// TwinCAT 3 PLC project TcoAteqMeasurementTests
// Title: TcoAteqMeasurementTests
// Company: Vortex.Library
// ProjectVersion: 0.6.0.913
// ProgramVersion: 3.1.4024.12
// libraries:
//   TcoAteqMeasurement, 0.6.0.913 (Vortex.Library)
//   Tc2_Standard, * (Beckhoff Automation GmbH)
//   Tc2_System, * (Beckhoff Automation GmbH)
//   Tc3_Module, * (Beckhoff Automation GmbH)
//   TcoIo, 0.6.0.913 (Vortex.Library)
//   TcoCore, 0.6.0.913 (Vortex.Library)
// project tree:
//   GVLs/ GVL.TcGVL
//   / PlcTask.TcTTO
//   POUs/ MAIN.TcPOU
//   Tests/TcoAteqG6/ eTcoAteqG6Tests.TcDUT, TcoAteqG6Simulator.TcPOU, TcoAteqG6TestContext.TcPOU
//   Tests/TcoContext/ WpfContext.TcPOU
// (motion and I/O tree: see PLC project tcoateqmeasurement)
// real-time tasks:
//   TASK PlcTask: cycle T#10ms, priority 20, ADS port 350
//   TASK PlcTask1: cycle T#10ms, priority 21, ADS port 351

CONFIGURATION TcoAteqMeasurementTests
    RESOURCE PLC ON TwinCAT3
        TASK PlcTask(INTERVAL := T#10ms, PRIORITY := 21);
        PROGRAM MAIN WITH PlcTask : MAIN;
    END_RESOURCE
END_CONFIGURATION

// ---- Tests/TcoAteqG6/eTcoAteqG6Tests.TcDUT
{attribute 'qualified_only'}
{attribute 'strict'}
TYPE eTcoAteqG6Tests :
(
	None := 0,
	Restore := 10,
	Run := 20,
	Reset := 30,
	SelectProgram := 40,
	StartCycle := 50,
	ReadLastResult := 60,
	SpecialCycle := 70,
	ReadParameters := 80,
	ReadPresetParameters := 90,
	ReadParameter := 100,
	InvokeStartCycle := 110,
	InvokeSelectProgram := 120,
	InvokeReset := 130
);
END_TYPE

// ---- GVLs/GVL.TcGVL
{attribute 'qualified_only'}
VAR_GLOBAL
	Ateq1 : TcoAteqMeasurement.TcoAteqG6Pn_IO_v_3_5_x;
END_VAR

// ---- POUs/MAIN.TcPOU
PROGRAM MAIN
VAR
	_g6TestContext : TcoAteqG6TestContext;

	_wpfContext : WpfContext;
	_wpfContextCall : BOOL := FALSE;
END_VAR

_g6TestContext.ProbeRun();

IF _wpfContextCall THEN
	_wpfContext.Run();
END_IF

END_PROGRAM

// ---- Tests/TcoAteqG6/TcoAteqG6TestContext.TcPOU
(*~
	<docu>
		<summary>
			Test context of TcoAteqG6Pn_v_3_5_x. _inImage is the input image of the instrument: written by the simulator
			when _simulate = TRUE, otherwise directly by the test. _outImage is what the component put on the wire.
		</summary>
	</docu>
~*)
FUNCTION_BLOCK TcoAteqG6TestContext EXTENDS TcoCore._internals_TcoContext
VAR
	_sut : TcoAteqMeasurement.TcoAteqG6Pn_v_3_5_x(THIS^);
	_io : TcoAteqMeasurement.TcoAteqG6Pn_IO_v_3_5_x;
	_sim : TcoAteqG6Simulator;
	_simulate : BOOL;
	_inImage : ARRAY[0..255] OF BYTE;
	_outImage : ARRAY[0..255] OF BYTE;
	_program : INT;
	_specialCycle : TcoAteqMeasurement.eTcoAteqG6_SpecialCycle_v_3_5_x;
	_instruction : BYTE;
	_parameter : TcoAteqMeasurement.eTcoAteqG6_ParameterId_v_3_5_x;
	_request : TcoAteqMeasurement.TcoAteqG6_ParameterRequest_v_3_5_x;
	_taskDone : BOOL;
	_taskError : BOOL;
	_startCycleBusy : BOOL;
	_selectProgramBusy : BOOL;
	_resetBusy : BOOL;
END_VAR
VAR
	{attribute 'hide'}
	_i : INT;
END_VAR

METHOD PROTECTED Main
//*************INSTRUMENT SIMULATOR*******
IF _simulate THEN
	_sim.Step(inoOut := _outImage, inoIn := _inImage);
END_IF

//*************INPUT IMAGE****************
MEMCPY(destAddr := ADR(_io.In.In1), srcAddr := ADR(_inImage[0]), n := 64);
MEMCPY(destAddr := ADR(_io.In.In2), srcAddr := ADR(_inImage[64]), n := 64);
MEMCPY(destAddr := ADR(_io.In.In3), srcAddr := ADR(_inImage[128]), n := 64);
MEMCPY(destAddr := ADR(_io.In.In4), srcAddr := ADR(_inImage[192]), n := 64);

CASE _testId OF
	eTcoAteqG6Tests.Restore:
		_sut.Restore();
		_sut._messenger.Clear();
		_sim.Reset();
		FOR _i := 0 TO 255 DO
			_inImage[_i] := 0;
		END_FOR
		_taskDone := FALSE;
		_taskError := FALSE;
		ProbeDoneWhen(TRUE);
	eTcoAteqG6Tests.Run:
		;
	eTcoAteqG6Tests.Reset:
		_taskDone := _sut.Reset().Done;
		_taskError := _sut.ResetTask.Error;
		ProbeDoneWhen(_taskDone OR _taskError);
	eTcoAteqG6Tests.SelectProgram:
		_taskDone := _sut.SelectProgram(_program).Done;
		_taskError := _sut.SelectProgramTask.Error;
		ProbeDoneWhen(_taskDone OR _taskError);
	eTcoAteqG6Tests.StartCycle:
		_taskDone := _sut.StartCycle(_program).Done;
		_taskError := _sut.StartCycleTask.Error;
		ProbeDoneWhen(_taskDone OR _taskError);
	eTcoAteqG6Tests.ReadLastResult:
		_taskDone := _sut.ReadLastResult().Done;
		_taskError := _sut.ReadLastResultTask.Error;
		ProbeDoneWhen(_taskDone OR _taskError);
	eTcoAteqG6Tests.SpecialCycle:
		_taskDone := _sut.SpecialCycle(_specialCycle, _instruction).Done;
		_taskError := _sut.SpecialCycleTask.Error;
		ProbeDoneWhen(_taskDone OR _taskError);
	eTcoAteqG6Tests.ReadParameters:
		_taskDone := _sut.ReadParameters(_request).Done;
		_taskError := _sut.ReadParametersTask.Error;
		ProbeDoneWhen(_taskDone OR _taskError);
	eTcoAteqG6Tests.ReadPresetParameters:
		_taskDone := _sut.ReadPresetParameters().Done;
		_taskError := _sut.ReadParametersTask.Error;
		ProbeDoneWhen(_taskDone OR _taskError);
	eTcoAteqG6Tests.ReadParameter:
		_taskDone := _sut.ReadParameter(_parameter).Done;
		_taskError := _sut.ReadParametersTask.Error;
		ProbeDoneWhen(_taskDone OR _taskError);
	eTcoAteqG6Tests.InvokeStartCycle:
		_sut.StartCycle(_program);
		ProbeDoneWhen(TRUE);
	eTcoAteqG6Tests.InvokeSelectProgram:
		_sut.SelectProgram(_program);
		ProbeDoneWhen(TRUE);
	eTcoAteqG6Tests.InvokeReset:
		_sut.Reset();
		ProbeDoneWhen(TRUE);
END_CASE

_sut(inoData := _io);

//*************OUTPUT IMAGE***************
MEMCPY(destAddr := ADR(_outImage[0]), srcAddr := ADR(_io.Out.Out1), n := 64);
MEMCPY(destAddr := ADR(_outImage[64]), srcAddr := ADR(_io.Out.Out2), n := 64);
MEMCPY(destAddr := ADR(_outImage[128]), srcAddr := ADR(_io.Out.Out3), n := 64);
MEMCPY(destAddr := ADR(_outImage[192]), srcAddr := ADR(_io.Out.Out4), n := 64);

_startCycleBusy := _sut.StartCycleTask.Busy;
_selectProgramBusy := _sut.SelectProgramTask.Busy;
_resetBusy := _sut.ResetTask.Busy;
END_METHOD

END_FUNCTION_BLOCK

// ---- Tests/TcoAteqG6/TcoAteqG6Simulator.TcPOU
(*~
	<docu>
		<summary>
			Simulated ATEQ G6 instrument (port of the AX FakeG6 harness). Each Step() plays one PLC cycle of the instrument
			against the output image: a rising command edge is echoed with error word FFFFh, the command completes after
			CommandCycles cycles (error word 0, or the command's own bit when it is in FailMask), the echo drops once the
			PLC drops the command bit. A started (special) cycle clears CycleEnd for CycleCycles cycles. Results are written
			into the input image exactly where the real instrument puts them.
		</summary>
	</docu>
~*)
FUNCTION_BLOCK TcoAteqG6Simulator
VAR
	// behaviour knobs
	CommandCycles : INT := 2;
	CycleCycles : INT := 3;
	FailMask : WORD;               // commands completing with an error
	SilentMask : WORD;             // commands never acknowledged
	StuckEchoMask : WORD;          // echo never released
	IgnoreProgramSelection : BOOL;
	NoCycle : BOOL;                // start accepted, cycle end never drops
	EndlessCycle : BOOL;           // cycle end never comes back
	ResultProgramOffset : INT;     // <> 0 -> stale last result
	ResultRelay : WORD := 16#0001;
	ResultAlarm : INT;
	// instrument state
	BusProgram : INT;              // 0-based, as on the bus
	CycleEnd : BOOL := TRUE;
	Echo : WORD;
	Error : WORD;
	// observations
	RisingEdges : INT;
	RaisedUnion : WORD;
	LastRaised : WORD;
	LastSpecialId : BYTE;
END_VAR
VAR
	_prev : WORD;
	_active : WORD;
	_busy : INT;
	_cycle : INT;
END_VAR

METHOD Reset
CommandCycles := 2;
CycleCycles := 3;
FailMask := 0;
SilentMask := 0;
StuckEchoMask := 0;
IgnoreProgramSelection := FALSE;
NoCycle := FALSE;
EndlessCycle := FALSE;
ResultProgramOffset := 0;
ResultRelay := 16#0001;
ResultAlarm := 0;
BusProgram := 0;
CycleEnd := TRUE;
Echo := 0;
Error := 0;
RisingEdges := 0;
RaisedUnion := 0;
LastRaised := 0;
LastSpecialId := 0;
_prev := 0;
_active := 0;
_busy := 0;
_cycle := 0;
END_METHOD

METHOD Step
VAR_IN_OUT
	inoOut : ARRAY[0..255] OF BYTE; // what the PLC put on the wire
	inoIn : ARRAY[0..255] OF BYTE;  // input image of the instrument
END_VAR
VAR
	cmd : WORD;
	rising : WORD;
	dropped : WORD;
END_VAR
cmd := TcoAteqMeasurement.TcoAteqG6_GetWord_v_3_5_x(inOffset := 16#00, inoImage := inoOut);
rising := cmd AND NOT _prev;
dropped := _prev AND NOT cmd;
IF rising <> 0 THEN
	RisingEdges := RisingEdges + 1;
	RaisedUnion := RaisedUnion OR rising;
	LastRaised := rising;
	IF (rising AND SilentMask) = 0 THEN
		_active := rising;
		Echo := Echo OR rising;
		Error := 16#FFFF;
		_busy := CommandCycles;
		IF (rising AND 16#0004) <> 0 THEN
			LastSpecialId := inoOut[16#08];
		END_IF
	END_IF
END_IF
IF _busy > 0 THEN
	_busy := _busy - 1;
	IF _busy = 0 THEN
		Complete(inoOut := inoOut, inoIn := inoIn);
	END_IF
END_IF
Echo := Echo AND NOT (dropped AND NOT StuckEchoMask);
IF _cycle > 0 AND NOT EndlessCycle THEN
	_cycle := _cycle - 1;
	IF _cycle = 0 THEN
		CycleEnd := TRUE;
		WriteLastResult(inoIn := inoIn);
	END_IF
END_IF
_prev := cmd;
WriteState(inoIn := inoIn);
END_METHOD

METHOD PRIVATE Complete
VAR_IN_OUT
	inoOut : ARRAY[0..255] OF BYTE;
	inoIn : ARRAY[0..255] OF BYTE;
END_VAR
IF (_active AND FailMask) <> 0 THEN
	Error := _active;
	RETURN;
END_IF
Error := 0;
IF _active = 16#0001 THEN
	CycleEnd := TRUE;
	_cycle := 0;
ELSIF _active = 16#0008 THEN
	IF NOT IgnoreProgramSelection THEN
		BusProgram := TcoAteqMeasurement.TcoAteqG6_GetInt_v_3_5_x(inOffset := 16#06, inoImage := inoOut);
	END_IF
ELSIF _active = 16#0002 OR _active = 16#0006 THEN
	IF NOT NoCycle THEN
		CycleEnd := FALSE;
		_cycle := CycleCycles;
	END_IF
ELSIF _active = 16#8000 THEN
	WriteLastResult(inoIn := inoIn);
ELSIF _active = 16#0020 THEN
	WriteParameters(inoOut := inoOut, inoIn := inoIn);
END_IF
END_METHOD

METHOD PRIVATE WriteState
VAR_IN_OUT
	inoIn : ARRAY[0..255] OF BYTE;
END_VAR
VAR
	status : WORD;
END_VAR
TcoAteqMeasurement.TcoAteqG6_SetWord_v_3_5_x(inOffset := 16#00, inValue := Echo, inoImage := inoIn);
TcoAteqMeasurement.TcoAteqG6_SetWord_v_3_5_x(inOffset := 16#02, inValue := Error, inoImage := inoIn);
TcoAteqMeasurement.TcoAteqG6_SetWord_v_3_5_x(inOffset := 16#06, inValue := INT_TO_WORD(BusProgram), inoImage := inoIn);
IF CycleEnd THEN
	status := 16#0020;
END_IF
TcoAteqMeasurement.TcoAteqG6_SetWord_v_3_5_x(inOffset := 16#0C, inValue := status, inoImage := inoIn);
END_METHOD

METHOD PRIVATE WriteLastResult
VAR_IN_OUT
	inoIn : ARRAY[0..255] OF BYTE;
END_VAR
TcoAteqMeasurement.TcoAteqG6_SetWord_v_3_5_x(inOffset := 16#20, inValue := INT_TO_WORD(BusProgram + ResultProgramOffset), inoImage := inoIn);
TcoAteqMeasurement.TcoAteqG6_SetWord_v_3_5_x(inOffset := 16#24, inValue := ResultRelay, inoImage := inoIn);
TcoAteqMeasurement.TcoAteqG6_SetWord_v_3_5_x(inOffset := 16#26, inValue := INT_TO_WORD(ResultAlarm), inoImage := inoIn);
TcoAteqMeasurement.TcoAteqG6_SetDint_v_3_5_x(inOffset := 16#28, inValue := 207000, inoImage := inoIn);
TcoAteqMeasurement.TcoAteqG6_SetDint_v_3_5_x(inOffset := 16#2C, inValue := 14000, inoImage := inoIn);
TcoAteqMeasurement.TcoAteqG6_SetDint_v_3_5_x(inOffset := 16#30, inValue := -108, inoImage := inoIn);
TcoAteqMeasurement.TcoAteqG6_SetDint_v_3_5_x(inOffset := 16#34, inValue := 1000, inoImage := inoIn);
END_METHOD

(*~
	<docu>
		<summary>
			Response value of every requested parameter = its identifier x 1000. The request (count + identifiers) is read from output 20h.
		</summary>
	</docu>
~*)
METHOD PRIVATE WriteParameters
VAR_IN_OUT
	inoOut : ARRAY[0..255] OF BYTE;
	inoIn : ARRAY[0..255] OF BYTE;
END_VAR
VAR
	i : INT;
	count : INT;
	id : WORD;
END_VAR
count := TcoAteqMeasurement.TcoAteqG6_GetInt_v_3_5_x(inOffset := 16#20, inoImage := inoOut);
FOR i := 0 TO count - 1 DO
	id := TcoAteqMeasurement.TcoAteqG6_GetWord_v_3_5_x(inOffset := 16#22 + 2 * i, inoImage := inoOut);
	TcoAteqMeasurement.TcoAteqG6_SetWord_v_3_5_x(inOffset := 16#20 + 6 * i, inValue := id, inoImage := inoIn);
	TcoAteqMeasurement.TcoAteqG6_SetDint_v_3_5_x(inOffset := 16#22 + 6 * i, inValue := WORD_TO_DINT(id) * 1000, inoImage := inoIn);
END_FOR
END_METHOD

END_FUNCTION_BLOCK

// ---- Tests/TcoContext/WpfContext.TcPOU
FUNCTION_BLOCK WpfContext EXTENDS TcoCore.TcoContext
VAR
	_serviceModeActive : BOOL;
	{attribute addProperty Name "<#ATEQ G6 PN#>"}
	_ateq1 : TcoAteqMeasurement.TcoAteqG6Pn_v_3_5_x(THIS^);
END_VAR

METHOD PROTECTED Main
IF _serviceModeActive THEN
	_ateq1.Service();
END_IF
_ateq1(inoData := GVL.Ateq1);
END_METHOD

END_FUNCTION_BLOCK
